// TwinCAT 3 PLC project PLCstudent
// ProgramVersion: 3.1.4026.20
// libraries:
//   Tc2_Standard, * (Beckhoff Automation GmbH)
//   Tc2_System, * (Beckhoff Automation GmbH)
// project tree:
//   GVLs/ GVL.TcGVL
//   / PlcTask.TcTTO
//   POUs/ FunktionBlockDiagram.TcPOU, MAIN.TcPOU, OUTPUT_TEXT.TcPOU, SPEED_CONTROL.TcPOU
// real-time tasks:
//   TASK PlcTask: cycle T#10ms, priority 20, ADS port 350
//   TASK PlcTask1: cycle T#10ms, priority 21, ADS port 351
// variable links:
//   PLCsim/PLCsim Instance <-> PLCstudent/PLCstudent Instance
//     PlcTask Inputs/GVL.isStatusText <-> PlcTask Outputs/GVL.qsStatusText
//     PlcTask Inputs/GVL.iwPumpSpeed <-> PlcTask Outputs/GVL.qwPumpSpeed
//     PlcTask Outputs/GVL.qwActualLevel <-> PlcTask Inputs/GVL.iwActualLevel

CONFIGURATION PLCstudent
    RESOURCE PLC ON TwinCAT3
        TASK PlcTask(INTERVAL := T#10ms, PRIORITY := 20);
        PROGRAM MAIN WITH PlcTask : MAIN;
    END_RESOURCE
END_CONFIGURATION

// ---- GVLs/GVL.TcGVL
{attribute 'qualified_only'}
VAR_GLOBAL

	qwPumpSpeed   		AT%Q* :  WORD; 	// Speed of the flow into the tank 0 - 100%
										// 40% slowly drain 50% stand still 60% filling
										

	qsStatusText 		AT%Q* : STRING := 'Test text'; // Text on the info display
	
	iwActualLevel 		AT%I* : WORD;  	// Level in the tank	
	
END_VAR

// ---- POUs/MAIN.TcPOU
PROGRAM MAIN
VAR
END_VAR


FunktionBlockDiagram();

END_PROGRAM

// ---- POUs/FunktionBlockDiagram.TcPOU
PROGRAM FunktionBlockDiagram
VAR
	ixLevel : INT;
	mxHighLevel : BOOL;
	mxLowerLevel : BOOL;
	mxLevel : INT;
	
	miProportional : INT := 10;
	miConst : INT := 50;
	miNewProp :  INT;
	
	msNormalLevel : STRING  := 'Normal Level';
	msHighLevel : STRING := 'High Level';
	msLowerLevel : STRING := 'Lower Level';
	
	
END_VAR

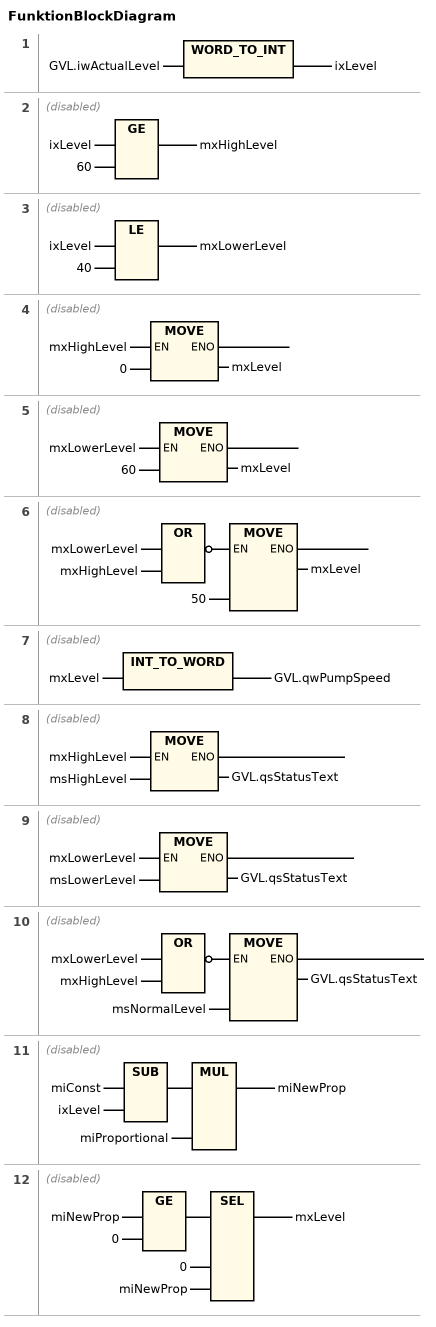
// NETWORK 1
ixLevel := WORD_TO_INT(GVL.iwActualLevel);

// NETWORK 2 (disabled)
// mxHighLevel := ixLevel >= 60;

// NETWORK 3 (disabled)
// mxLowerLevel := ixLevel <= 40;

// NETWORK 4 (disabled)
// IF mxHighLevel THEN mxLevel := 0; END_IF

// NETWORK 5 (disabled)
// IF mxLowerLevel THEN mxLevel := 60; END_IF

// NETWORK 6 (disabled)
// IF NOT (mxLowerLevel OR mxHighLevel) THEN mxLevel := 50; END_IF

// NETWORK 7 (disabled)
// GVL.qwPumpSpeed := INT_TO_WORD(mxLevel);

// NETWORK 8 (disabled)
// IF mxHighLevel THEN GVL.qsStatusText := msHighLevel; END_IF

// NETWORK 9 (disabled)
// IF mxLowerLevel THEN GVL.qsStatusText := msLowerLevel; END_IF

// NETWORK 10 (disabled)
// IF NOT (mxLowerLevel OR mxHighLevel) THEN GVL.qsStatusText := msNormalLevel; END_IF

// NETWORK 11 (disabled)
// miNewProp := (miConst - ixLevel) * miProportional;

// NETWORK 12 (disabled)
// mxLevel := SEL(miNewProp >= 0, 0, miNewProp);

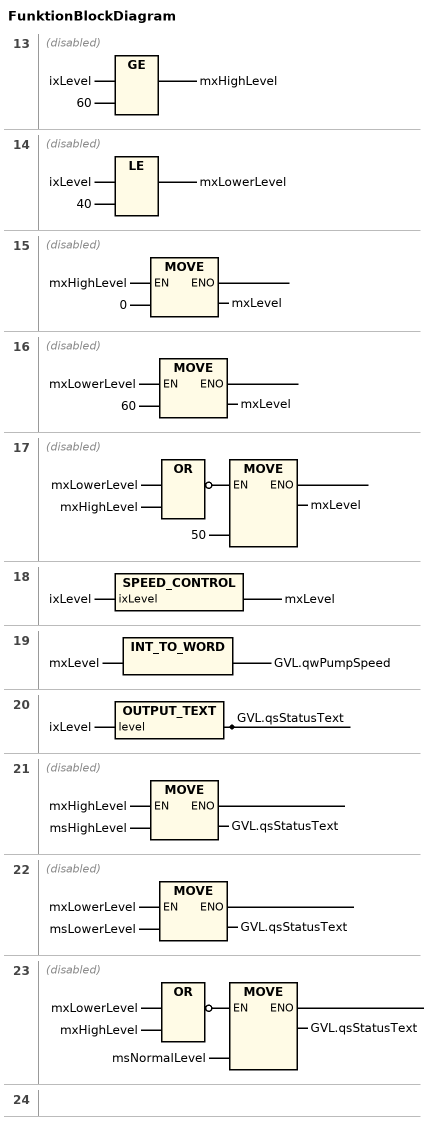
// NETWORK 13 (disabled)
// mxHighLevel := ixLevel >= 60;

// NETWORK 14 (disabled)
// mxLowerLevel := ixLevel <= 40;

// NETWORK 15 (disabled)
// IF mxHighLevel THEN mxLevel := 0; END_IF

// NETWORK 16 (disabled)
// IF mxLowerLevel THEN mxLevel := 60; END_IF

// NETWORK 17 (disabled)
// IF NOT (mxLowerLevel OR mxHighLevel) THEN mxLevel := 50; END_IF

// NETWORK 18
mxLevel := SPEED_CONTROL(ixLevel := ixLevel);

// NETWORK 19
GVL.qwPumpSpeed := INT_TO_WORD(mxLevel);

// NETWORK 20
GVL.qsStatusText := OUTPUT_TEXT(level := ixLevel);

// NETWORK 21 (disabled)
// IF mxHighLevel THEN GVL.qsStatusText := msHighLevel; END_IF

// NETWORK 22 (disabled)
// IF mxLowerLevel THEN GVL.qsStatusText := msLowerLevel; END_IF

// NETWORK 23 (disabled)
// IF NOT (mxLowerLevel OR mxHighLevel) THEN GVL.qsStatusText := msNormalLevel; END_IF

// NETWORK 24

END_PROGRAM

// ---- POUs/SPEED_CONTROL.TcPOU
FUNCTION SPEED_CONTROL : INT
VAR_INPUT
	ixLevel : INT;
END_VAR

SPEED_CONTROL := (50 - ixLevel) * 10;
IF SPEED_CONTROL < 0 THEN;
	SPEED_CONTROL := 0;
END_IF

END_FUNCTION

// ---- POUs/OUTPUT_TEXT.TcPOU
FUNCTION OUTPUT_TEXT : STRING
VAR_INPUT
	level : INT;
END_VAR
VAR
END_VAR

IF level >= 60 THEN;
	OUTPUT_TEXT := 'High Level';
ELSIF level <= 40 THEN;
	OUTPUT_TEXT := 'Low Level';
ELSE
	OUTPUT_TEXT := 'Normal Level';
END_IF

END_FUNCTION
